FUNCTION_BLOCK Filling
VAR_INPUT
	diEnabled : BOOL;
END_VAR
VAR_OUTPUT
	doEnabled : BOOL;
END_VAR
VAR_IN_OUT
	FillingPhase : TPhaseFilling;
	FillingValve : TValve;
END_VAR
VAR
END_VAR

{region "REGION Aut/Man"}
    // switching state of engine - automatic or manual control (default state is manual)
  	IF FillingPhase.Cmd.ManCtrl THEN
      	FillingPhase.State.ManCtrl := TRUE;
		FillingPhase.State.AutCtrl := FALSE;
	ELSIF FillingPhase.Cmd.AutCtrl THEN
        FillingPhase.State.ManCtrl := FALSE;
		FillingPhase.State.AutCtrl := TRUE; 
    END_IF;
		 
	IF (NOT FillingPhase.State.AutCtrl AND NOT FillingPhase.State.ManCtrl) THEN
		FillingPhase.State.ManCtrl := TRUE;
	END_IF

	FillingPhase.Cmd.ManCtrl := FALSE;
	FillingPhase.Cmd.AutCtrl := FALSE;
{endregion}

{region "ManCtrl"}
    // processing manual actions - if command is processed, it is sets to FALSE even if can't be processed
    // Phase commands are start, stop, pause and resume 
    // Start - open filling valve 
    // Stop - close filling valve
    // Pause - close filling valve
    // Resume - open filling valve
    // real states of phase are wrote into states in phase structure
    IF FillingPhase.State.ManCtrl THEN
		IF FillingPhase.State.Idle AND FillingPhase.Cmd.StartMan THEN
			FillingPhase.State.Running := TRUE;
			FillingPhase.State.Idle := FALSE;
			FillingPhase.State.Paused := FALSE;
		 	FillingPhase.State.Done := FALSE;
		ELSIF FillingPhase.Cmd.StopMan THEN
			FillingPhase.State.Running := FALSE;
			FillingPhase.State.Idle := TRUE;
			FillingPhase.State.Paused := FALSE;
		ELSIF FillingPhase.State.Running AND FillingPhase.Cmd.PauseMan THEN
			FillingPhase.State.Running := FALSE;
			FillingPhase.State.Idle := FALSE;
			FillingPhase.State.Paused := TRUE;
		ELSIF FillingPhase.State.Paused AND FillingPhase.Cmd.ResumeMan THEN
			FillingPhase.State.Running := TRUE;
			FillingPhase.State.Idle := FALSE;
			FillingPhase.State.Paused := FALSE;
			FillingPhase.State.Done := FALSE;
		END_IF
    END_IF;
	
	FillingPhase.Cmd.StartMan := FALSE;
	FillingPhase.Cmd.StopMan := FALSE;
	FillingPhase.Cmd.PauseMan := FALSE;
	FillingPhase.Cmd.ResumeMan := FALSE;
{endregion}

{region "AutCtrl"}
    // if request to run in automatic mode and phase can be run in automatic mode switch phase to running
    IF FillingPhase.State.AutCtrl THEN
		IF FillingPhase.State.Idle AND FillingPhase.Cmd.StartAut THEN
			FillingPhase.State.Running := TRUE;
			FillingPhase.State.Idle := FALSE;
		 	FillingPhase.State.Done := FALSE;
		ELSIF FillingPhase.Cmd.StopAut THEN
			FillingPhase.State.Running := FALSE;
			FillingPhase.State.Idle := TRUE;
			FillingPhase.State.Paused := FALSE;
		END_IF
    END_IF;
	
	FillingPhase.Cmd.StartAut := FALSE;
	FillingPhase.Cmd.StopAut := FALSE;
{endregion}

{region "Done"}
    //every phase should have finish condition - filling phase - if water level is above requested level
    //after that done state should be set to 1
    IF FillingPhase.State.Running AND (FillingPhase.WaterLevel >= FillingPhase.ParamFillLevel - 0.083) THEN // edit based on speed of simulation 
        FillingPhase.Cmd.StopMan := TRUE;
        FillingPhase.Cmd.StopAut := TRUE;
        FillingPhase.State.Done := TRUE;
    END_IF;

    IF FillingPhase.Cmd.ResetDone THEN
        FillingPhase.State.Done := FALSE;
        FillingPhase.Cmd.ResetDone := FALSE;
    END_IF;
{endregion}

{region "States"}
	//Command valve in cases of states
    IF FillingPhase.State.Running THEN
        FillingValve.Cmd.Req2OpenAut := TRUE;
        FillingValve.Cmd.Req2CloseAut := FALSE;
    ELSE
        FillingValve.Cmd.Req2OpenAut := FALSE;
        FillingValve.Cmd.Req2CloseAut := TRUE;
    END_IF;
{endregion}


// delault state of phase - if not any state sets state to idle
IF NOT FillingPhase.State.Idle AND NOT FillingPhase.State.Paused AND NOT FillingPhase.State.Running THEN
    FillingPhase.State.Idle := 1;
END_IF;

// write binary states into int value for visualization
IF FillingPhase.State.Idle THEN
    FillingPhase.State.Stateint := Global.PhIdle;
ELSIF FillingPhase.State.Running THEN
    FillingPhase.State.Stateint := Global.PhRunning;
ELSE
    FillingPhase.State.Stateint := Global.PhPause;
END_IF;

// Ponechte pro moznost retezeni volani bloku v LAD
doEnabled := diEnabled;

END_FUNCTION_BLOCK

(* stored: Version 1.1.0.1, ProductVersion 3.1.4026.21
   POU Filling: Id {9d4dcb01-ad56-4326-9456-8cd473ff054e}, SpecialFunc None *)
